{attribute 'qualified_only'}
{attribute 'strict'}
TYPE E_Filling_Mode :
(
	Not_Selected := 0,
	Bin,
	Bin_Cyrculation,
	Line_Cyrculation
	
);
END_TYPE

(* stored: Version 1.1.0.1, ProductVersion 3.1.4024.15
   DUT E_Filling_Mode: Id {19fb8745-ab6c-486c-9bac-aa81ae860b52} *)
